// TIA Portal V21 export
// export: Created 2026-11-18T10:00:00.0000000Z, ExportSetting None
FUNCTION_BLOCK "FB_Station"   // FB20, LAD
{ S7_Optimized_Access := 'TRUE' }
// stored: MemoryReserve 100, SetENOAutomatically false
   VAR_INPUT
      Enable : Bool;
      Init : Bool;
   END_VAR
   VAR_OUTPUT
      Lamp : Bool;
   END_VAR
   VAR
      Seq : "FB_Sequence";
      Run : Bool;
      Fault : Bool;   // set after 5 s
      T_Fault : TON_TIME;
   END_VAR
BEGIN

REGION Network 1: Sequence
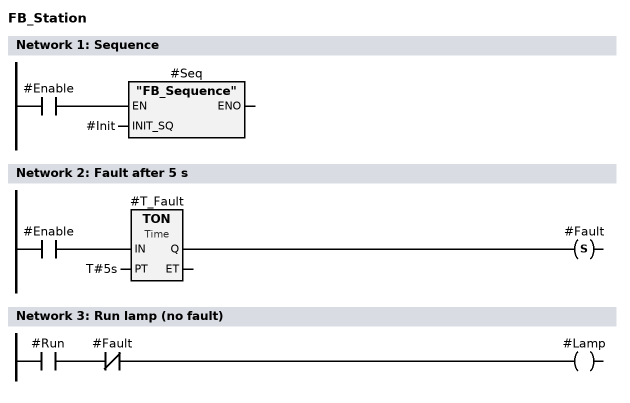
   RUNG wire#powerrail
      Contact( #Enable )
      #Seq(INIT_SQ := #Init)
   END_RUNG
   // the same network as SCL:
   IF #Enable THEN
       #Seq(INIT_SQ := #Init);   // "FB_Sequence"
   END_IF;
END_REGION

REGION Network 2: Fault after 5 s
   RUNG wire#powerrail
      Contact( #Enable )
      { S7_Templates := "time_type := Time" } #T_Fault.TON(pt := T#5s, et =>)
      S_Coil( #Fault )
   END_RUNG
   // the same network as SCL:
   #T_Fault(IN := #Enable, PT := T#5s);   // TON
   IF #T_Fault.Q THEN #Fault := TRUE; END_IF;
END_REGION

REGION Network 3: Run lamp (no fault)
   RUNG wire#powerrail
      Contact( #Run )
      I_Contact( #Fault )
      Coil( #Lamp )
   END_RUNG
   // the same network as SCL:
   #Lamp := #Run AND NOT #Fault;
END_REGION
END_FUNCTION_BLOCK
